// LS Electric XG5000 project: day3last
// PLC LSPLC

PROGRAM NewProgram (task: 스캔 프로그램)

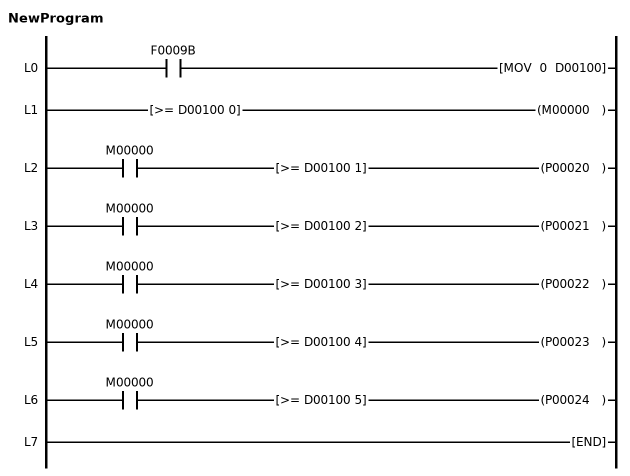
; L0
LOAD      F0009B
MOV       0 D00100
; L1
LOAD>=    D00100 0
OUT       M00000
; L2
LOAD      M00000
AND>=     D00100 1
OUT       P00020
; L3
LOAD      M00000
AND>=     D00100 2
OUT       P00021
; L4
LOAD      M00000
AND>=     D00100 3
OUT       P00022
; L5
LOAD      M00000
AND>=     D00100 4
OUT       P00023
; L6
LOAD      M00000
AND>=     D00100 5
OUT       P00024
; L7
END